// TIA Portal V20 export
// export: Created 2026-10-12T05:42:35.5976794Z, ExportSetting WithDefaults, DisplayName Totally Integrated Automation Portal, DisplayVersion V20, DisplayName TIA Portal Openness, DisplayVersion V20, DisplayName TIA Portal Teamcenter Gateway, DisplayVersion V20, DisplayName TIA Portal Version Control Interface, DisplayVersion V20, DisplayName SINAMICS Startdrive Advanced, DisplayVersion V20 SP1 Update 2, DisplayName SINAMICS Startdrive G110M, G120, G120C, G120D, G120P, G115D, DisplayVersion V20 SP1 Update 2, DisplayName SINAMICS Startdrive G130, G150, S120, S150, SINAMICS MV, G220, S200, S210, DisplayVersion V20 SP1 Update 2, DisplayName STEP 7 Professional, DisplayVersion V20, DisplayName STEP 7 Safety, DisplayVersion V20, DisplayName WinCC Basic/Comfort/Advanced, DisplayVersion V20, DisplayName WinCC Professional, DisplayVersion V20, DisplayName WinCC Unified, DisplayVersion V20
FUNCTION_BLOCK "FB_PressDemoRelease"   // FB5, SCL
{ S7_Optimized_Access := 'TRUE' }
VERSION : 0.1
// stored: AutoNumber true, IsIECCheckEnabled false, IsRetainMemResEnabled false, MemoryReserve 100, SetENOAutomatically false, UDAEnableTagReadback false
   VAR_INPUT
      AirPressureOk : Bool;
      DoorClosed : Bool;
      DoorHealthy : Bool;
      RamHealthy : Bool;
      SlideHealthy : Bool;
      SlideInside : Bool;
      TwoHandHeld : Bool;
   END_VAR
   VAR
      Conditions { ExternalWritable := 'False'; S7_SetPoint := 'True'} : "ST_PressDemoReleaseConditions";
      ModeStart { ExternalWritable := 'False'; S7_SetPoint := 'True'} : "FRK_PermCtx";
      RamExtend { ExternalWritable := 'False'; S7_SetPoint := 'True'} : "FRK_PermCtx";
   END_VAR
BEGIN

   #Conditions.ModeStartAirPressureOk := #AirPressureOk;
   #Conditions.RamGuardClosed := #DoorClosed;
   #Conditions.RamSlideInside := #SlideInside;
   #Conditions.RamDevicesHealthy := #RamHealthy AND #DoorHealthy AND #SlideHealthy;
   #Conditions.RamAirPressureOk := #AirPressureOk;
   #Conditions.RamTwoHandHeld := #TwoHandHeld;
   "FRK_PermBegin"(Perm := #ModeStart);
   "FRK_PermCondition"(Perm := #ModeStart,
                       Label := 'project.condition.ModeStartAirPressureOk',
                       Ok := #Conditions.ModeStartAirPressureOk);
   "FRK_PermBegin"(Perm := #RamExtend);
   "FRK_PermCondition"(Perm := #RamExtend,
                       Label := 'project.condition.RamGuardClosed',
                       Ok := #Conditions.RamGuardClosed);
   "FRK_PermCondition"(Perm := #RamExtend,
                       Label := 'project.condition.RamSlideInside',
                       Ok := #Conditions.RamSlideInside);
   "FRK_PermCondition"(Perm := #RamExtend,
                       Label := 'project.condition.RamDevicesHealthy',
                       Ok := #Conditions.RamDevicesHealthy);
   "FRK_PermCondition"(Perm := #RamExtend,
                       Label := 'project.condition.RamAirPressureOk',
                       Ok := #Conditions.RamAirPressureOk);
   "FRK_PermCondition"(Perm := #RamExtend,
                       Label := 'project.condition.RamTwoHandHeld',
                       Ok := #Conditions.RamTwoHandHeld);
END_FUNCTION_BLOCK
